(* IEC 61131-3 sources: RootPLC/bench/tasks/latch-start-stop/reference, 1 file *)

(* ---- solution.st ---- *)
PROGRAM PRG_Motor
VAR_INPUT
    start, stop : BOOL;
END_VAR
VAR_OUTPUT
    running : BOOL;
END_VAR
running := (start OR running) AND NOT stop;
END_PROGRAM
